// Generated by voz_llm_plc_agent
// Target: Siemens TIA Portal V18 - SCL external source
// Review and compile before any download to physical hardware.

FUNCTION_BLOCK "PLC_PRG"
{ S7_Optimized_Access := 'TRUE' }
VERSION : 0.1
VAR_INPUT
   I_Start : Bool := FALSE;
   I_Stop : Bool := FALSE;
   I_Emergency : Bool := FALSE;
END_VAR
VAR_OUTPUT
   Q_Contactor_Principal : Bool := FALSE;
END_VAR
VAR
   M_Contactor_RunLatch : Bool;
   M_Contactor_PrincipalLatch : Bool;
   M_Contactor_RunLatch_StartPrevious : Bool;
   M_Contactor_RunLatch_StartInitialized : Bool;
   M_Contactor_RunLatch_StartPulse : Bool;
END_VAR
BEGIN
#M_Contactor_RunLatch_StartPulse := #M_Contactor_RunLatch_StartInitialized AND #I_Start AND NOT #M_Contactor_RunLatch_StartPrevious;
#M_Contactor_RunLatch_StartPrevious := #I_Start;
#M_Contactor_RunLatch_StartInitialized := TRUE;
(* Enclavamiento de motor con prioridad de paro y emergencia *)
IF #I_Emergency OR #I_Stop THEN
    #M_Contactor_RunLatch := FALSE;
ELSIF #M_Contactor_RunLatch_StartPulse THEN
    #M_Contactor_RunLatch := TRUE;
END_IF;

#Q_Contactor_Principal := #M_Contactor_RunLatch AND NOT #I_Emergency;
END_FUNCTION_BLOCK

DATA_BLOCK "DB_PLC_PRG"
{ S7_Optimized_Access := 'TRUE' }
VERSION : 0.1
NON_RETAIN
"PLC_PRG"
BEGIN
END_DATA_BLOCK

ORGANIZATION_BLOCK "Main"
{ S7_Optimized_Access := 'TRUE' }
VERSION : 0.1
BEGIN
   "DB_PLC_PRG"(
      I_Start := "I_Start",
      I_Stop := "I_Stop",
      I_Emergency := "I_Emergency",
      Q_Contactor_Principal => "Q_Contactor_Principal"
   );
END_ORGANIZATION_BLOCK
